// TIA Portal V21 export
// export: Created 2026-10-23T20:43:14.6549864Z, ExportSetting WithDefaults, DisplayName Totally Integrated Automation Portal, DisplayVersion V21 Update 1, DisplayName SINAMICS Startdrive Advanced, DisplayVersion V21 HF2, DisplayName SINAMICS Startdrive G110M, G120, G120C, G120D, G120P, G115D, DisplayVersion V21 HF2, DisplayName SINAMICS Startdrive G130, G150, S120, S150, G200, G220, S200, S210, S220, Innomotics MVD, DisplayVersion V21 HF2, DisplayName STEP 7 Professional, DisplayVersion V21 Update 1, DisplayName STEP 7 Safety, DisplayVersion V21, DisplayName Tech WebApplication, DisplayVersion V21, DisplayName WinCC Basic/Comfort/Advanced, DisplayVersion V21 Update 1, DisplayName WinCC Unified, DisplayVersion V21 Update 1
FUNCTION "FC_AnaTempRead" : Int   // FC10, SCL
TITLE = Analyzer: Temp read before written
{ S7_Optimized_Access := 'TRUE' }
VERSION : 0.1
// Rule C26c: Sum is read before it is written
// stored: AutoNumber true, IsIECCheckEnabled false, SetENOAutomatically false, UDAEnableTagReadback false
   VAR_INPUT
      Value : Int;   // Value to add
   END_VAR
   VAR_TEMP
      Sum : Int;   // Temporary sum
   END_VAR
BEGIN

       #Sum := #Sum + #Value;
       #FC_AnaTempRead := #Sum;
END_FUNCTION
